// TIA Portal V20 export
// export: Created 2026-10-20T12:40:08.6583016Z, ExportSetting WithDefaults, DisplayName Totally Integrated Automation Portal, DisplayVersion V20 Update 6, DisplayName TIA Portal Openness, DisplayVersion V20 Update 6, DisplayName TIA Portal Version Control Interface, DisplayVersion V20 Update 6, DisplayName SINAMICS Startdrive Advanced, DisplayVersion V20 SP1, DisplayName SINAMICS Startdrive G130, G150, S120, S150, SINAMICS MV, G220, S200, S210, DisplayVersion V20 SP1, DisplayName SINAMICS Startdrive G110M, G120, G120C, G120D, G120P, G115D, DisplayVersion V20 SP1, DisplayName STEP 7 Professional, DisplayVersion V20 Update 6, DisplayName STEP 7 Safety, DisplayVersion V20 Update 2, DisplayName WinCC Basic/Comfort/Advanced, DisplayVersion V20 Update 6, DisplayName WinCC Unified, DisplayVersion V20 Update 6
DATA_BLOCK "SICK_AFx60_Data_DB"   // DB120
{ S7_Optimized_Access := 'TRUE' }
VERSION : 0.1
// stored: AutoNumber true, DBAccessibleFromOPCUA true, IsOnlyStoredInLoadMemory false, IsRetainMemResEnabled false, IsWriteProtectedInAS false, MemoryReserve 100
   VAR
      "Absolute Encoder 1" { S7_SetPoint := 'True'} : "ST_SICK_AFx60";
      "Absolute Encoder 2" { S7_SetPoint := 'True'} : "ST_SICK_AFx60";
      "Absolute Encoder 3" { S7_SetPoint := 'True'} : "ST_SICK_AFx60";
      "Absolute Encoder 4" { S7_SetPoint := 'True'} : "ST_SICK_AFx60";
      "Absolute Encoder 5" { S7_SetPoint := 'True'} : "ST_SICK_AFx60";
   END_VAR
BEGIN
END_DATA_BLOCK
